// TIA Portal V21 export
// export: Created 2026-10-26T12:54:42.3373989Z, ExportSetting WithDefaults, DisplayName Totally Integrated Automation Portal, DisplayVersion V21 Update 3, DisplayName TIA Portal Test Suite Advanced, DisplayVersion V21 Update 1, DisplayName SINAMICS Startdrive Advanced, DisplayVersion V21 Update 1, DisplayName SINAMICS Startdrive G130, G150, S120, S150, G200, G210, G210C, G210X, G220, S200, S210, S220, Innomotics MVD, DisplayVersion V21 Update 1, DisplayName SINAMICS Startdrive G110M, G120, G120C, G120D, G120P, G115D, DisplayVersion V21 Update 1, DisplayName STEP 7 Professional, DisplayVersion V21 Update 3, DisplayName STEP 7 Safety, DisplayVersion V21, DisplayName Tech WebApplication, DisplayVersion V21, DisplayName WinCC Basic/Comfort/Advanced, DisplayVersion V21 Update 3, DisplayName WinCC Professional, DisplayVersion V21 Update 3, DisplayName WinCC Unified, DisplayVersion V21 Update 3
FUNCTION_BLOCK "TgpUnit_IecEffect"   // FB2, SCL
VERSION : 0.1
// stored: Access Unpublished, AutoNumber true, IsIECCheckEnabled false, IsRetainMemResEnabled false, MemoryReserve 100, Namespace TiaMcp_UnitA, SetENOAutomatically false, UDAEnableTagReadback false
   VAR_INPUT
      Enable : Bool;
   END_VAR
   VAR_OUTPUT
      Active : Bool;
   END_VAR
   VAR
      RetainedMarker : Int := 17;
      Timer_TON { S7_SetPoint := 'True'} : TON_TIME;
      Timer_TOF { S7_SetPoint := 'True'} : TOF_TIME;
      Timer_TP { S7_SetPoint := 'True'} : TP_TIME;
      Counter_CTU { S7_SetPoint := 'True'} : CTU_INT;
      Counter_CTD { S7_SetPoint := 'True'} : CTD_INT;
      Counter_CTUD { S7_SetPoint := 'True'} : CTUD_INT;
   END_VAR
BEGIN

    #Active := #Enable;
END_FUNCTION_BLOCK
